{attribute 'qualified_only' := ''}
{attribute 'strict' := ''}
TYPE E_PointType :
(
	POINTTYPE_XY := 1,
	POINTTYPE_XYVA := 2
);
END_TYPE

(* stored: Version 1.1.0.1, ProductVersion 3.1.4024.12
   DUT E_PointType: Id {5a9f2a88-4c97-4e5d-8749-f736d636a191} *)
